(* Logix 5000 project; controller DSFW_0512_C_FCB_S1_SPN vendor 1 type 14 code 77 rev 20.12; software revision 20.06; part 3 of 3 *)
(* tags used below, declared in another part *)
   Compressor_Superheat : REAL;
   EEV_101_Auto_Manual : BOOL;
   EEV_101_Manual_Output : REAL;
   EEV_101_Pressure_Setpoint : REAL;
   EEV_101_Run_PIDE : BOOL;
   EEV_101_Run_Temp_PIDE : BOOL;
   EEV_101_Stop_PIDE : BOOL;
   EEV_101_Superheat_Setpoint : REAL;
   EEV_102_Auto_Manual : BOOL;
   EEV_102_Manual_Output : REAL;
   EEV_102_SH_Setpoint : REAL;
   EEV_102_Stop_PIDE : BOOL;
   Evaporator_Superheat : REAL;
   PT_101_Reactor_Supply_Pressure : REAL;
   PT_102_Compressor_Suction_Pressure : REAL;
   PT_102_Offset : REAL;
   PT_103_Compressor_Discharge_Pressure : REAL;
   PT_103_Offset : REAL;
   PT_104_Evaporator_Suction_Pressure : REAL;
   PT_104_Offset : REAL;
   Reactor_Batch_CV_as_SP : REAL;
   Reactor_Batch_PID_Start : BOOL;
   Reactor_Batch_PID_Stop : BOOL;
   Reactor_Batch_PV : REAL;
   TCV_101_Auto_Manual : BOOL;
   TCV_101_Manual_Output : REAL;
   TCV_101_Run_PIDE : BOOL;
   TCV_101_Stop_PIDE : BOOL;
   TE_101_Liquid_Line_Temperature : REAL;
   TE_101_Offset : REAL;
   TE_102_Evaporator_Suction_Temperature : REAL;
   TE_102_Offset : REAL;
   TE_103_Compressor_Suction_Temperature : REAL;
   TE_103_Offset : REAL;
   TE_105_Reactor_Supply_Temperature : REAL;
   Temperature_Setpoint : REAL;
(* Refrigeration_Control, continued *)

ROUTINE Sensors   (* ladder *)
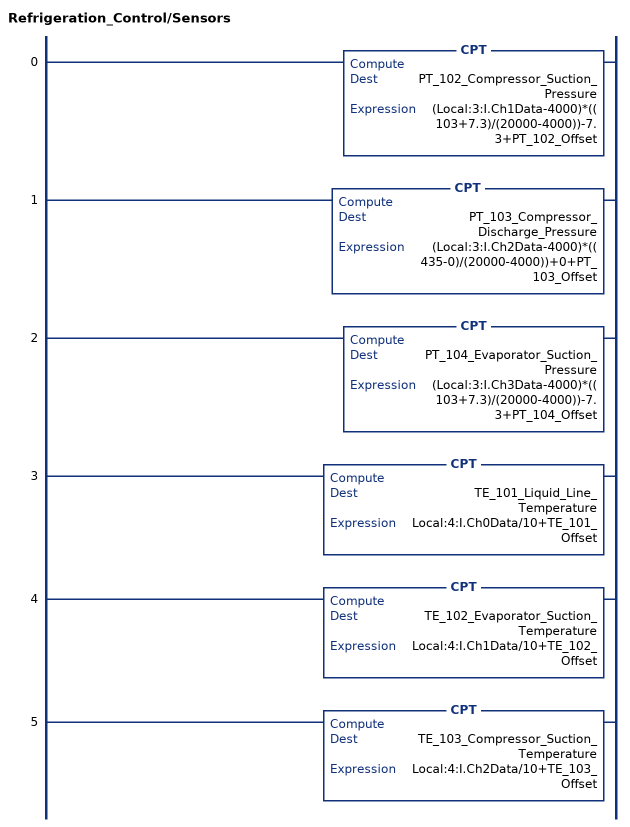
   0: CPT(PT_102_Compressor_Suction_Pressure,(Local:3:I.Ch1Data-4000)*((103+7.3)/(20000-4000))-7.3+PT_102_Offset);
   1: CPT(PT_103_Compressor_Discharge_Pressure,(Local:3:I.Ch2Data-4000)*((435-0)/(20000-4000))+0+PT_103_Offset);
   2: CPT(PT_104_Evaporator_Suction_Pressure,(Local:3:I.Ch3Data-4000)*((103+7.3)/(20000-4000))-7.3+PT_104_Offset);
   3: CPT(TE_101_Liquid_Line_Temperature,Local:4:I.Ch0Data/10+TE_101_Offset);
   4: CPT(TE_102_Evaporator_Suction_Temperature,Local:4:I.Ch1Data/10+TE_102_Offset);
   5: CPT(TE_103_Compressor_Suction_Temperature,Local:4:I.Ch2Data/10+TE_103_Offset);
END_ROUTINE
END_PROGRAM

PROGRAM Refrigeration_PID_Calculations   (* main routine TCV_101 *)
VAR
   BOR_01 : FBD_BOOLEAN_OR;
   BOR_02 : FBD_BOOLEAN_OR;
   BOR_03 : FBD_BOOLEAN_OR;
   BOR_04 : FBD_BOOLEAN_OR := (In2 := 1, Out := 1);
   ESEL_01 : SELECT_ENHANCED := (InsUsed := 3, SelectorMode := 2, OperSelector := 1, ProgProgReq := 1, SelectedIn := 1, ProgOper := 1);
   ESEL_02 : SELECT_ENHANCED := (InsUsed := 1, SelectorMode := 2);
   PIDE_01 : PID_ENHANCED := (PV := 40.73446, PVEUMax := 100.0, SPProg := 12.0, SPOper := 12.0, SPHLimit := 100.0, RatioProg := 1.0, RatioOper := 1.0, RatioHLimit := 1.0, RatioLLimit := 1.0, CVProg := 43.558277, CVOper := 43.558277, CVEUMax := 20000.0, CVEUMin := 4000.0, CVHLimit := 100.0, CVLLimit := 8.0, ControlAction := 1, PGain := 9.0, IGain := 1.9, PVEDerivative := 1, DSmoothing := 1, PVHHLimit := 150.0, PVHLimit := 100.0, PVLLimit := 2.0, PVLLLimit := 1.0, ProgValueReset := 1, RTSTime := 1, CVEU := 10969.324, CV := 43.558277, SP := 12.0, SPPercent := 12.0, PVPercent := 40.73446, E := 28.734459, EPercent := 28.734459, InitPrimary := 1, Ratio := 1.0, Auto := 1, DeltaT := 0.2);
   PIDE_02 : PID_ENHANCED := (PV := 40.73446, PVEUMax := 100.0, SPProg := 12.0, SPOper := 12.0, SPHLimit := 100.0, RatioProg := 1.0, RatioOper := 1.0, RatioHLimit := 1.0, RatioLLimit := 1.0, CVProg := 43.558277, CVOper := 43.558277, CVEUMax := 20000.0, CVEUMin := 4000.0, CVHLimit := 100.0, CVLLimit := 8.0, ControlAction := 1, PGain := 9.0, IGain := 1.9, PVEDerivative := 1, DSmoothing := 1, PVHHLimit := 150.0, PVHLimit := 100.0, PVLLimit := 2.0, PVLLLimit := 1.0, ProgValueReset := 1, RTSTime := 1, CVEU := 10969.324, CV := 43.558277, SP := 12.0, SPPercent := 12.0, PVPercent := 40.73446, E := 28.734459, EPercent := 28.734459, InitPrimary := 1, Ratio := 1.0, Auto := 1, DeltaT := 0.2);
   PIDE_03 : PID_ENHANCED := (PV := 40.73446, PVEUMax := 100.0, SPProg := 12.0, SPOper := 12.0, SPHLimit := 100.0, RatioProg := 1.0, RatioOper := 1.0, RatioHLimit := 1.0, RatioLLimit := 1.0, CVProg := 43.558277, CVOper := 43.558277, CVEUMax := 20000.0, CVEUMin := 4000.0, CVHLimit := 100.0, CVLLimit := 8.0, ControlAction := 1, PGain := 9.0, IGain := 1.9, PVEDerivative := 1, DSmoothing := 1, PVHHLimit := 150.0, PVHLimit := 100.0, PVLLimit := 2.0, PVLLLimit := 1.0, ProgValueReset := 1, RTSTime := 1, CVEU := 10969.324, CV := 43.558277, SP := 12.0, SPPercent := 12.0, PVPercent := 40.73446, E := 28.734459, EPercent := 28.734459, InitPrimary := 1, Ratio := 1.0, Auto := 1, DeltaT := 0.2);
   PIDE_04 : PID_ENHANCED := (PV := 40.73446, PVEUMax := 100.0, SPProg := 12.0, SPOper := 12.0, SPHLimit := 100.0, RatioProg := 1.0, RatioOper := 1.0, RatioHLimit := 1.0, RatioLLimit := 1.0, CVProg := 43.558277, CVOper := 43.558277, CVEUMax := 20000.0, CVEUMin := 4000.0, CVHLimit := 100.0, CVLLimit := 8.0, ControlAction := 1, PGain := 9.0, IGain := 1.9, PVEDerivative := 1, DSmoothing := 1, PVHHLimit := 150.0, PVHLimit := 100.0, PVLLimit := 2.0, PVLLLimit := 1.0, ProgValueReset := 1, RTSTime := 1, CVEU := 10969.324, CV := 43.558277, SP := 12.0, SPPercent := 12.0, PVPercent := 40.73446, E := 28.734459, EPercent := 28.734459, InitPrimary := 1, Ratio := 1.0, Auto := 1, DeltaT := 0.2);
   PIDE_05 : PID_ENHANCED := (PV := 40.73446, PVEUMax := 100.0, SPProg := 12.0, SPOper := 12.0, SPHLimit := 100.0, RatioProg := 1.0, RatioOper := 1.0, RatioHLimit := 1.0, RatioLLimit := 1.0, CVProg := 43.558277, CVOper := 43.558277, CVEUMax := 20000.0, CVEUMin := 4000.0, CVHLimit := 100.0, CVLLimit := 8.0, ControlAction := 1, PGain := 9.0, IGain := 1.9, PVEDerivative := 1, DSmoothing := 1, PVHHLimit := 150.0, PVHLimit := 100.0, PVLLimit := 2.0, PVLLLimit := 1.0, ProgValueReset := 1, RTSTime := 1, CVEU := 10969.324, CV := 43.558277, SP := 12.0, SPPercent := 12.0, PVPercent := 40.73446, E := 28.734459, EPercent := 28.734459, InitPrimary := 1, Ratio := 1.0, Auto := 1, DeltaT := 0.2);
   PIDE_06 : PID_ENHANCED := (PV := 40.73446, PVEUMax := 100.0, SPProg := 12.0, SPOper := 12.0, SPHLimit := 100.0, RatioProg := 1.0, RatioOper := 1.0, RatioHLimit := 1.0, RatioLLimit := 1.0, CVProg := 43.558277, CVOper := 43.558277, CVEUMax := 20000.0, CVEUMin := 4000.0, CVHLimit := 100.0, CVLLimit := 8.0, ControlAction := 1, PGain := 9.0, IGain := 1.9, PVEDerivative := 1, DSmoothing := 1, PVHHLimit := 150.0, PVHLimit := 100.0, PVLLimit := 2.0, PVLLLimit := 1.0, ProgValueReset := 1, RTSTime := 1, CVEU := 10969.324, CV := 43.558277, SP := 12.0, SPPercent := 12.0, PVPercent := 40.73446, E := 28.734459, EPercent := 28.734459, InitPrimary := 1, Ratio := 1.0, Auto := 1, DeltaT := 0.2);
   SEL_01 : SELECT := (In1 := 20.0, In2 := 18.941616, SelectorIn := 1, Out := 18.941616);
END_VAR

ROUTINE EEV_101   (* function block diagram *)
   SHEET 1
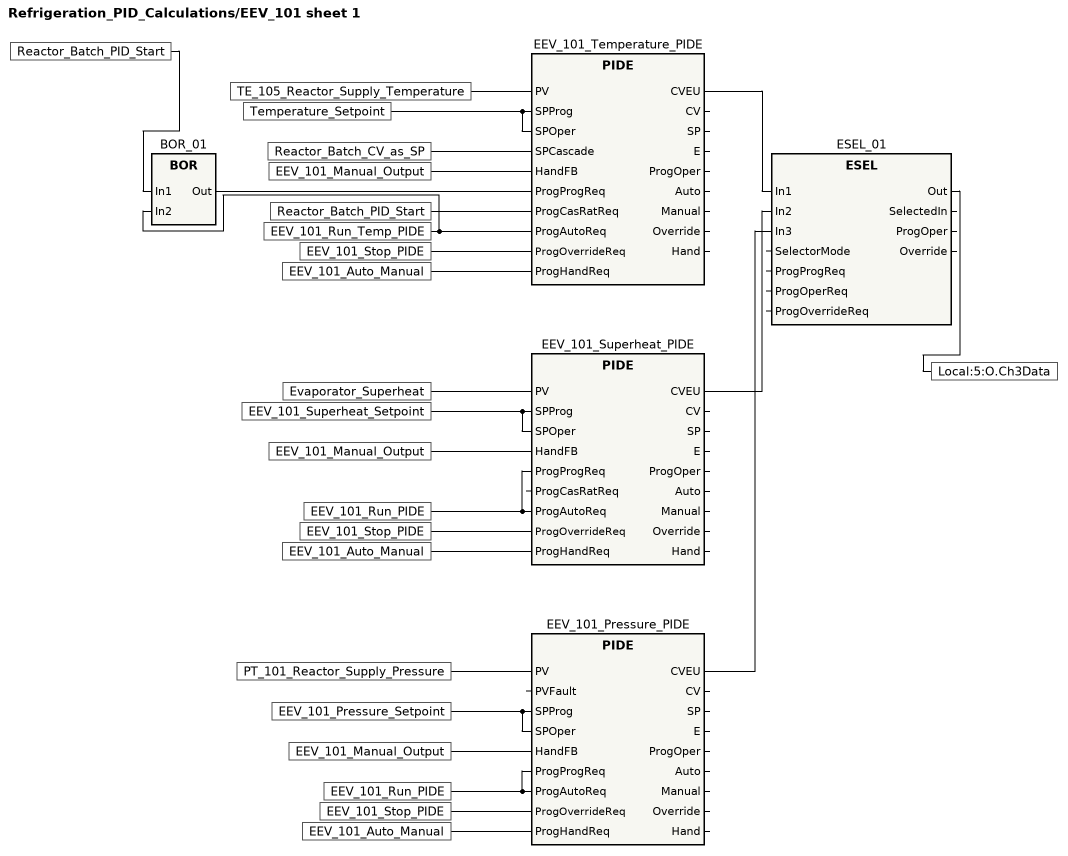
   BOR_01 : BOR(In1 := Reactor_Batch_PID_Start, In2 := EEV_101_Run_Temp_PIDE);
   EEV_101_Temperature_PIDE : PIDE(PV := TE_105_Reactor_Supply_Temperature, SPProg := Temperature_Setpoint, SPOper := Temperature_Setpoint, SPCascade := Reactor_Batch_CV_as_SP, HandFB := EEV_101_Manual_Output, ProgProgReq := BOR_01.Out, ProgCasRatReq := Reactor_Batch_PID_Start, ProgAutoReq := EEV_101_Run_Temp_PIDE, ProgOverrideReq := EEV_101_Stop_PIDE, ProgHandReq := EEV_101_Auto_Manual);   // unwired pins: CV SP E ProgOper Auto Manual Override Hand
   EEV_101_Superheat_PIDE : PIDE(PV := Evaporator_Superheat, SPProg := EEV_101_Superheat_Setpoint, SPOper := EEV_101_Superheat_Setpoint, HandFB := EEV_101_Manual_Output, ProgProgReq := EEV_101_Run_PIDE, ProgAutoReq := EEV_101_Run_PIDE, ProgOverrideReq := EEV_101_Stop_PIDE, ProgHandReq := EEV_101_Auto_Manual);   // unwired pins: ProgCasRatReq CV SP E ProgOper Auto Manual Override Hand
   EEV_101_Pressure_PIDE : PIDE(PV := PT_101_Reactor_Supply_Pressure, SPProg := EEV_101_Pressure_Setpoint, SPOper := EEV_101_Pressure_Setpoint, HandFB := EEV_101_Manual_Output, ProgProgReq := EEV_101_Run_PIDE, ProgAutoReq := EEV_101_Run_PIDE, ProgOverrideReq := EEV_101_Stop_PIDE, ProgHandReq := EEV_101_Auto_Manual);   // unwired pins: PVFault CV SP E ProgOper Auto Manual Override Hand
   ESEL_01 : ESEL(In1 := EEV_101_Temperature_PIDE.CVEU, In2 := EEV_101_Superheat_PIDE.CVEU, In3 := EEV_101_Pressure_PIDE.CVEU);   // unwired pins: SelectorMode ProgProgReq ProgOperReq ProgOverrideReq SelectedIn ProgOper Override
   Local:5:O.Ch3Data := ESEL_01.Out;
END_ROUTINE

ROUTINE EEV_102   (* function block diagram *)
   SHEET 1
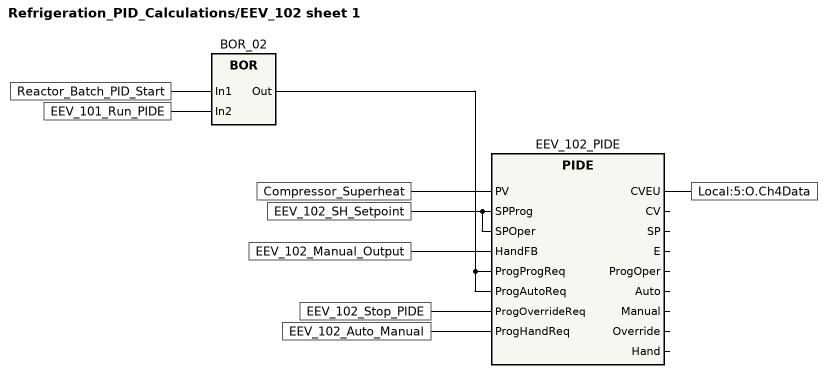
   BOR_02 : BOR(In1 := Reactor_Batch_PID_Start, In2 := EEV_101_Run_PIDE);
   EEV_102_PIDE : PIDE(PV := Compressor_Superheat, SPProg := EEV_102_SH_Setpoint, SPOper := EEV_102_SH_Setpoint, HandFB := EEV_102_Manual_Output, ProgProgReq := BOR_02.Out, ProgAutoReq := BOR_02.Out, ProgOverrideReq := EEV_102_Stop_PIDE, ProgHandReq := EEV_102_Auto_Manual);   // unwired pins: CV SP E ProgOper Auto Manual Override Hand
   Local:5:O.Ch4Data := EEV_102_PIDE.CVEU;
END_ROUTINE

ROUTINE TCV_101   (* function block diagram *)
   SHEET 1
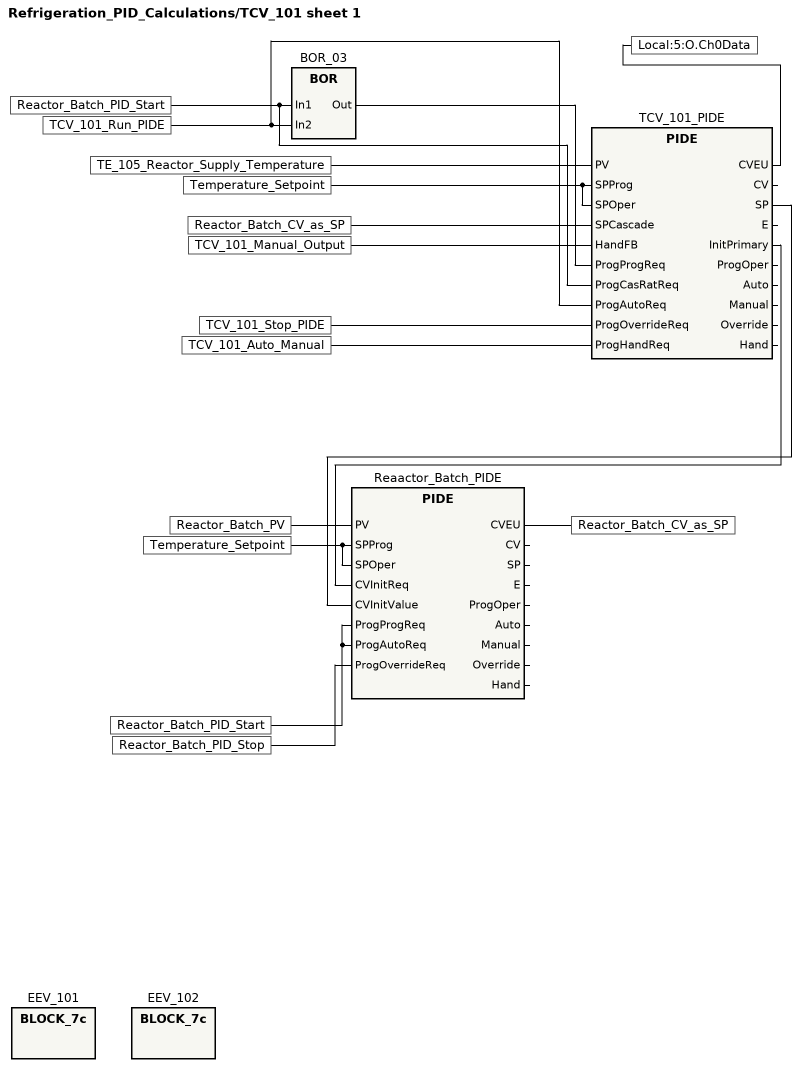
   EEV_101 : BLOCK_7c();
   EEV_102 : BLOCK_7c();
   BOR_03 : BOR(In1 := Reactor_Batch_PID_Start, In2 := TCV_101_Run_PIDE);
   TCV_101_PIDE : PIDE(PV := TE_105_Reactor_Supply_Temperature, SPProg := Temperature_Setpoint, SPOper := Temperature_Setpoint, SPCascade := Reactor_Batch_CV_as_SP, HandFB := TCV_101_Manual_Output, ProgProgReq := BOR_03.Out, ProgCasRatReq := Reactor_Batch_PID_Start, ProgAutoReq := TCV_101_Run_PIDE, ProgOverrideReq := TCV_101_Stop_PIDE, ProgHandReq := TCV_101_Auto_Manual);   // unwired pins: CV E ProgOper Auto Manual Override Hand
   Reaactor_Batch_PIDE : PIDE(PV := Reactor_Batch_PV, SPProg := Temperature_Setpoint, SPOper := Temperature_Setpoint, CVInitReq := TCV_101_PIDE.InitPrimary, CVInitValue := TCV_101_PIDE.SP, ProgProgReq := Reactor_Batch_PID_Start, ProgAutoReq := Reactor_Batch_PID_Start, ProgOverrideReq := Reactor_Batch_PID_Stop);   // unwired pins: CV SP E ProgOper Auto Manual Override Hand
   Reactor_Batch_CV_as_SP := Reaactor_Batch_PIDE.CVEU;
   Local:5:O.Ch0Data := TCV_101_PIDE.CVEU;
END_ROUTINE
END_PROGRAM
